(* IEC 61131-3 sources: beedance/examples/unit_tests, 4 files *)

(* ---- motor.st ---- *)
(* The code under test: a motor starter and a scaling function.
   The tests are in motor_tests.st; run them with
       beedance -test motor.st motor_tests.st *)

TYPE MotorStatus :
STRUCT
    running : BOOL;  (* the motor is running *)
    starts  : INT;   (* how many times it started *)
END_STRUCT;
END_TYPE

(* Scale converts a raw analog input (0..27648) to percent (0..100). *)
FUNCTION Scale : REAL
VAR_INPUT raw : INT; END_VAR
Scale := INT_TO_REAL(raw) * 100.0 / 27648.0;
END_FUNCTION

(* MotorStarter runs the motor once start has been held for delay, and
   stops it at once on stop or fault. *)
FUNCTION_BLOCK MotorStarter
VAR_INPUT
    start : BOOL;
    stop  : BOOL;
    fault : BOOL;
    delay : TIME;
END_VAR
VAR_OUTPUT
    run    : BOOL;
    status : MotorStatus;
END_VAR
VAR
    startDelay : TON;
END_VAR
startDelay(IN := start AND NOT stop AND NOT fault, PT := delay);
IF startDelay.Q AND NOT run THEN
    run := TRUE;
    status.starts := status.starts + 1;
END_IF;
IF stop OR fault THEN
    run := FALSE;
END_IF;
status.running := run;
END_FUNCTION_BLOCK

(* ---- failing.st ---- *)
(* Tests that fail on purpose, to show how each kind of failure is
   reported. Run with
       beedance -test -engines all -go-timeout 5s motor.st failing.st *)

(* A failed check: failures <> 0, with the message of the last one. *)
PROGRAM TEST_WrongExpectation
VAR_OUTPUT failures : INT; message : STRING; END_VAR
IF ABS(Scale(raw := 27648) - 99.0) > 0.001 THEN
    failures := failures + 1; message := 'expected 99 %';
END_IF;
END_PROGRAM

(* Never done: a test with done that is not done after -max-scans fails. *)
PROGRAM TEST_NeverDone
VAR_OUTPUT failures : INT; done : BOOL; END_VAR
VAR m : MotorStarter; END_VAR
m(start := TRUE, stop := TRUE, delay := T#1s);  (* stop holds it off *)
done := m.run;
END_PROGRAM

(* A runaway loop: the evaluator and the VM stop it with their per-scan
   budget; the go engine stops its process after -go-timeout. *)
PROGRAM TEST_RunawayLoop
VAR_OUTPUT failures : INT; END_VAR
VAR i : INT; END_VAR
WHILE TRUE DO
    i := i + 1;
END_WHILE;
END_PROGRAM

(* Not a test by the convention: it has no VAR_OUTPUT failures. *)
PROGRAM TEST_NoFailuresOutput
VAR x : INT; END_VAR
x := 1;
END_PROGRAM

(* ---- motor_tests.st ---- *)
(* Unit tests for motor.st. Every PROGRAM named TEST_... is a test:

     VAR_OUTPUT failures : INT;    checks that failed: 0 to pass
     VAR_OUTPUT message  : STRING; optional: what failed
     VAR_OUTPUT done     : BOOL;   optional: run scan by scan until TRUE

   Without done a test runs one scan. With done it runs scan by scan on a
   simulated clock (-interval apart, 10 ms by default) until done is TRUE. *)

(* One scan: a function's results. *)
PROGRAM TEST_Scale
VAR_OUTPUT failures : INT; message : STRING; END_VAR
IF ABS(Scale(raw := 0)) > 0.001 THEN
    failures := failures + 1; message := 'Scale(0) <> 0';
END_IF;
IF ABS(Scale(raw := 27648) - 100.0) > 0.001 THEN
    failures := failures + 1; message := 'Scale(27648) <> 100';
END_IF;
IF ABS(Scale(raw := 13824) - 50.0) > 0.001 THEN
    failures := failures + 1; message := 'Scale(13824) <> 50';
END_IF;
END_PROGRAM

(* Scan by scan: the motor must not run before its 5 s delay, and must
   run once it has passed. *)
PROGRAM TEST_MotorStartsAfterDelay
VAR_OUTPUT failures : INT; message : STRING; done : BOOL; END_VAR
VAR
    m     : MotorStarter;
    scans : INT;
END_VAR
scans := scans + 1;
m(start := TRUE, stop := FALSE, fault := FALSE, delay := T#5s);
(* At 10 ms a scan, scan 400 is at 3.99 s: too early to run. *)
IF scans = 400 AND m.run THEN
    failures := failures + 1; message := 'ran before the delay';
END_IF;
IF m.run THEN
    IF m.status.starts <> 1 THEN
        failures := failures + 1; message := 'starts <> 1';
    END_IF;
    done := TRUE;
END_IF;
END_PROGRAM

(* A sequence of steps: start, run, then a fault stops the motor at once. *)
PROGRAM TEST_MotorStopsOnFault
VAR_OUTPUT failures : INT; message : STRING; done : BOOL; END_VAR
VAR
    m     : MotorStarter;
    scans : INT;
    fault : BOOL;
END_VAR
scans := scans + 1;
fault := scans >= 20;  (* the fault comes at scan 20 *)
m(start := TRUE, stop := FALSE, fault := fault, delay := T#100ms);
IF scans = 19 AND NOT m.run THEN
    failures := failures + 1; message := 'not running before the fault';
END_IF;
IF scans = 20 THEN
    IF m.run OR m.status.running THEN
        failures := failures + 1; message := 'still running on fault';
    END_IF;
    done := TRUE;
END_IF;
END_PROGRAM

(* A long timer: a 5-minute delay takes 30,001 scans at the default 10 ms,
   301 with -interval 1s. The clock is simulated, so it runs in well under
   a second per engine, not 5 minutes. *)
PROGRAM TEST_LongDelay
VAR_OUTPUT failures : INT; message : STRING; done : BOOL; END_VAR
VAR m : MotorStarter; END_VAR
m(start := TRUE, delay := T#5m);
done := m.run;
END_PROGRAM

(* ---- precision.st ---- *)
(* REAL precision differs between engines: the evaluator and the VM hold a
   REAL in 64 bits, transpiled Go in 32 (iec.REAL is a float32), so 100/3
   is 33.333333 on one and 33.333332 on the other. -tol is the relative
   tolerance for comparing REAL and LREAL values between engines:

       beedance -test -engines all motor.st precision.st            agree
       beedance -test -engines all -tol 1e-9 motor.st precision.st  DIFFER *)

PROGRAM TEST_RealPrecision
VAR_OUTPUT failures : INT; END_VAR
VAR third : REAL; END_VAR
third := Scale(raw := 9216);  (* 9216 / 27648 * 100 = 33.33... *)
IF ABS(third - 33.3333) > 0.001 THEN
    failures := failures + 1;
END_IF;
END_PROGRAM
